// Mitsubishi GX Works2 project: test1   PLC: FX3U/FX3UC

PROGRAM MAIN
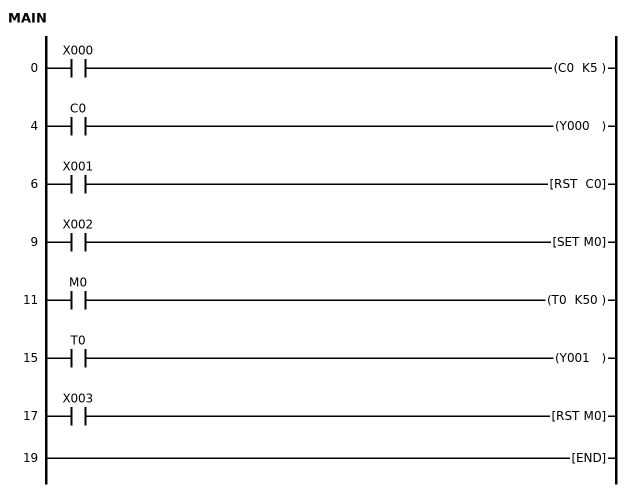
0     LD      X000
      OUT     C0 K5
4     LD      C0
      OUT     Y000
6     LD      X001
      RST     C0
9     LD      X002
      SET     M0
11    LD      M0
      OUT     T0 K50
15    LD      T0
      OUT     Y001
17    LD      X003
      RST     M0
19    END
END_PROGRAM
